(*
SPDX-FileCopyrightText: c 2026 Oleksandr Tiutyk <trofimich@gmail.com>
SPDX-License-Identifier: MIT
License: https://opensource.org/license/mit
*)

(*!
<summary>Checks assigning an empty builder to a populated target without allocating a builder buffer.</summary>
<description>
Uses one task and stays at a stable address while assertions are bound to this instance.
</description>
*)

{attribute 'no_assign'}
{attribute 'no_explicit_call' := 'do not call this function block directly'}
FUNCTION_BLOCK WideStringBuilderEmptyTest EXTENDS TOF_Testing.SingleCycleTest
VAR_STAT
	{attribute 'hide'}
	_ClassName : STRING := __POUNAME();
END_VAR
VAR
	_Builder : TOF_Core.WideStringBuilder;
END_VAR

(*!
<summary>Checks assigning an empty builder to a populated target without allocating a builder buffer.</summary>
<description>
The builder is persistent so teardown can release its buffer after an unexpected hook exception.
</description>
*)
METHOD PROTECTED ExecuteTest
VAR
	target : WSTRING := "previous contents";
	copied : BOOL;
END_VAR
copied := _Builder.AssignToString(targetString := target);
Assert.ThatBool(
	actual := copied AND_THEN target = "",
	message := "Assigning an empty builder must clear the target and succeed"
).IsTrue();
Assert.ThatBool(
	actual := _Builder.StringLength = 0 AND_THEN _Builder.Capacity = 0,
	message := "Assigning an empty builder must leave it unallocated"
).IsTrue();
END_METHOD

(*!
<summary>Releases the builder buffer before reporting the case result.</summary>
<description>
Safe after partial initialization and after explicit cleanup in the scenario.
</description>
*)
METHOD PROTECTED AfterTest
_Builder.Clear(releaseMemory := TRUE);
END_METHOD

//! <summary>Borrows the concrete class name. Callers must not modify it.</summary>
{attribute 'monitoring' := 'call'}
PROPERTY ClassName : REFERENCE TO STRING
GET
ClassName REF= _ClassName;
END_GET
END_PROPERTY

//! <summary>Borrows the compiler-initialized namespace name. Callers must not modify it.</summary>
{attribute 'monitoring' := 'call'}
PROPERTY NamespaceName : REFERENCE TO STRING
GET
NamespaceName REF= CurrentNamespace.Name;
END_GET
END_PROPERTY

//! <summary>Reports the concrete instance size in bytes.</summary>
{attribute 'monitoring' := 'call'}
PROPERTY SelfSize : ULINT
GET
SelfSize := XSIZEOF(THIS^);
END_GET
END_PROPERTY

END_FUNCTION_BLOCK

(* stored: Version 1.1.0.1
   POU WideStringBuilderEmptyTest: Id {82aecb06-8ab5-44af-b642-55f9dc49cbf2}, SpecialFunc None
   Method ExecuteTest: Id {49c26210-0a95-4753-905e-e7279cfab967}
   Method AfterTest: Id {7a3a04a2-fc4c-407c-a8fd-49570c8ccfdd}
   Property ClassName: Id {778f1200-8c33-4975-a5d7-c2da8f5ecbd8}
   Get Get: Id {b77dbbc3-17f2-4d48-a926-3cb4f16b645b}
   Property NamespaceName: Id {69773380-1189-4125-9cfe-86165603e5f0}
   Get Get: Id {d7e8ea10-b298-4dea-8010-b332be474c5a}
   Property SelfSize: Id {b2cefdd4-7c20-4777-a7f7-87f62dd988be}
   Get Get: Id {3c3470bd-e790-40e3-ab0c-06026ab06d10} *)
